// TIA Portal V20 export
// export: Created 2026-10-19T18:41:49.54429Z, ExportSetting WithDefaults, DisplayName Totally Integrated Automation Portal, DisplayVersion V20 Update 6, DisplayName TIA Portal Openness, DisplayVersion V20 Update 6, DisplayName TIA Portal Version Control Interface, DisplayVersion V20 Update 6, DisplayName SINAMICS Startdrive Advanced, DisplayVersion V20 SP1, DisplayName SINAMICS Startdrive G130, G150, S120, S150, SINAMICS MV, G220, S200, S210, DisplayVersion V20 SP1, DisplayName SINAMICS Startdrive G110M, G120, G120C, G120D, G120P, G115D, DisplayVersion V20 SP1, DisplayName STEP 7 Professional, DisplayVersion V20 Update 6, DisplayName STEP 7 Safety, DisplayVersion V20 Update 2, DisplayName WinCC Basic/Comfort/Advanced, DisplayVersion V20 Update 6, DisplayName WinCC Unified, DisplayVersion V20 Update 6
DATA_BLOCK "Barcode_FB_DB_1"   // DB144
VERSION : 0.1
// stored: AutoNumber true, DBAccessibleFromOPCUA true, InstanceOfName Barcode_Station_FB, InstanceOfType FB
"Barcode_Station_FB"
   // VAR_INPUT
   //    Sick_Result : String;
   // END_VAR
   // VAR_OUTPUT
   //    "Counter" : UInt;
   // END_VAR
   // VAR_IN_OUT
   //    Station_Control : "Barcode_Station_UDT";
   //    Auto_Start_Lector : Bool;
   //    Auto_Stop_Lector : Bool;
   // END_VAR
   // VAR
   //    State : UInt;
   //    R_Start_DB { S7_SetPoint := 'True'} : R_TRIG;
   //    T_Read_DB { S7_SetPoint := 'True'} : TON_TIME;
   // END_VAR
BEGIN
END_DATA_BLOCK
